(* IEC 61131-3 sources: codesys-framework/txt/application/WeVe Core (library)/10 Mode/Events, 2 files *)

(* ---- E_ModeEvents.dut.st ---- *)
// Events van de mode-laag (FB_ModeService en alle FB_Mode's). Index in FB_ModeEventGroup, niet de event-ID.
// Geen 'strict': de waarden worden als INT doorgegeven aan de EventGroup.
{attribute 'qualified_only'}
TYPE E_ModeEvents :
(
	// FB_ModeService
	ModeRequest := 0,
	ModeRequestInvalid,

	// FB_Mode
	StartRequestInvalid,
	ResetRequestInvalid,
	UserRequestInvalid,

	Count				// altijd laatste
);
END_TYPE

(* ---- FB_ModeEventGroup.pou.st ---- *)
// Events van de mode-laag. Eén instantie, gedeeld door FB_ModeService en alle FB_Mode's.
// Bevat enkel eenmalige meldingen (Log): er is geen toestand die modes met elkaar delen.
// De mode staat in de boodschap via %0.
//   fbModeEvents : FB_ModeEventGroup(fbLogger := fbLogger, nSubMachine := 0, nSubMachineId := 0);
FUNCTION_BLOCK FB_ModeEventGroup EXTENDS FB_EventGroup
VAR_INPUT
END_VAR
VAR_OUTPUT
END_VAR
VAR
	_afbEvents 		: ARRAY[0..E_ModeEvents.Count] OF FB_Event;		// slot Count blijft ongebruikt
END_VAR

// --- BEGIN IMPLEMENTATION ---
